// LS Electric XG5000 project: NewPLC
// PLC LSPLC
// module base 0 slot 0: 입력 모듈:XGI-D21A (DC 24V 입력, 8점 (전류소스/싱크입력))
// module base 0 slot 1: 입력 모듈:XGI-D22A/B (DC 24V 입력, 16점 (전류소스 싱크공용/ 전류소스 입력))
// module base 0 slot 2: 입력 모듈:XGI-D24A/B (DC 24V 입력, 32점 (전류소스 싱크공용/ 전류소스 입력))
// module base 0 slot 3: 입력 모듈:XGI-D28A/B (DC 24V 입력, 64점 (전류소스 싱크공용/ 전류소스 입력))
// module base 0 slot 4: 입력 모듈:XGI-A12A (AC 110V 입력, 16점)
// module base 0 slot 5: 입력 모듈:XGI-A21A/C (AC 220V 입력, 8점(8점/COM) / 8점(1점/COM))
// module base 0 slot 6: 입력 모듈:XGI-D21D (진단기능 내장형 DC24V 입력, 8점)
// module base 0 slot 7: 입출력 모듈:XGH-DT4A (DC 24V 입력, 트랜지스터 출력 32점 )
// module base 0 slot 8: 전용 모듈:XGI-LBDA (AC 110V 램프 단선검출 입력, 6점)
// module base 0 slot 9: 전용 모듈:XGI-LBDB (AC/DC 10V 램프 단선검출 입력, 6점)
// module base 0 slot 10: FDEnet:XGL-EDMT (전용 Ethernet 통신 모듈, 전기 Master)
// module base 0 slot 11: FDEnet:XGL-EDMF (전용 Ethernet 통신 모듈, 광 Master)
// module base 1 slot 0: 출력 모듈:XGQ-RY1A (릴레이 출력, 8점 (2A용, 단독 COM.))
// module base 1 slot 1: 출력 모듈:XGQ-RY2A/B (릴레이 출력, 16점 (2A용, Varistor 없음/Varistor 부착))
// module base 1 slot 2: 출력 모듈:XGQ-TR1C (트랜지스터 출력, 8점 (2A용, 싱크출력))
// module base 1 slot 3: 출력 모듈:XGQ-TR2A/B (트랜지스터 출력, 16점 (0.5A용, 싱크출력/소스출력))
// module base 1 slot 4: 출력 모듈:XGQ-TR4A/B (트랜지스터 출력, 32점 (0.1A용, 싱크출력/소스출력))
// module base 1 slot 5: 출력 모듈:XGQ-TR8A/B (트랜지스터 출력, 64점 (0.1A용, 싱크출력/소스출력))
// module base 1 slot 6: 출력 모듈:XGQ-SS2A (트라이액 출력, 16점 (1A용))
// module base 1 slot 7: 출력 모듈:XGQ-RY1D (진단기능 내장형 Relay 출력, 8점)
// module base 1 slot 8: 고속카운터 모듈:XGF-HO2A (고속카운터 펄스(OC) 입력형, 2채널)
// module base 1 slot 9: 고속카운터 모듈:XGF-HD2A (고속카운터 펄스(LD) 입력형, 2채널)
// module base 1 slot 10: 고속카운터 모듈:XGF-HO8A (고속카운터 펄스(OC) 입력형, 8채널)
// module base 1 slot 11: Dnet:XGL-DMEA/B (Dnet 통신 모듈, DeviceNet Master)
// module base 2 slot 0: 아날로그입력 모듈:XGF-AV8A (A/D 전압 입력형 8채널)
// module base 2 slot 1: 아날로그입력 모듈:XGF-AC8A (A/D 전류 입력형 8채널)
// module base 2 slot 2: 아날로그입력 모듈:XGF-AD4S (A/D 절연형 4채널)
// module base 2 slot 3: 아날로그입력 모듈:XGF-AD8A (A/D 전압/전류 입력형 8채널)
// module base 2 slot 4: 아날로그입력 모듈:XGF-AD16A (A/D 전압/전류 입력형 16채널)
// module base 2 slot 5: 아날로그입력 모듈:XGF-AC4H (HART 인터페이스 아날로그 전류입력, 4채널)
// module base 2 slot 6: 아날로그입력 모듈:XGF-AW4S (A/D 절연형 4채널(2선 입력형))
// module base 2 slot 7: 모션제어 모듈:XGF-M16M (모션 전용네트 (M-II)형, 16축)
// module base 2 slot 8: 모션제어 모듈:XGF-M32E (네트워크 표준형, 32축)
// module base 2 slot 9: 데이터로그 모듈:XGF-DL16A (데이터 로그 모듈)
// module base 2 slot 10: SOE모듈:XGF-SOEA (이벤트 기록 모듈)
// module base 2 slot 11: Rnet:XGL-RMEA/B (Rnet 통신 모듈, Rnet Master)
// module base 3 slot 0: 아날로그출력 모듈:XGF-DV4A (D/A 전압 출력형 4채널)
// module base 3 slot 1: 아날로그출력 모듈:XGF-DV8A (D/A 전압 출력형 8채널)
// module base 3 slot 2: 아날로그출력 모듈:XGF-DC4A (D/A 전류 출력형 4채널)
// module base 3 slot 3: 아날로그출력 모듈:XGF-DC8A (D/A 전류 출력형 8채널)
// module base 3 slot 4: 아날로그출력 모듈:XGF-DV4S (D/A 절연형 4채널(전압형))
// module base 3 slot 5: 아날로그출력 모듈:XGF-DC4S (D/A 절연형 4채널(전류형))
// module base 3 slot 6: 아날로그출력 모듈:XGF-DC4H (HART 인터페이스 아날로그 전류출력, 4채널)
// module base 3 slot 7: 아날로그출력 모듈:XGF-DA4S (D/A 절연형, 4채널)
// module base 3 slot 8: 온도입력 모듈:XGF-RD4A (온도 입력형 4채널)
// module base 3 slot 9: 온도입력 모듈:XGF-RD4S (온도 입력형 4채널(절연형))
// module base 3 slot 10: 온도입력 모듈:XGF-TC4S (온도 입력형 (절연형 4채널))
// module base 3 slot 11: 온도입력 모듈:XGF-RD8A (측온저항체 센서 입력형 8채널)

PROGRAM NewProgram (task: 스캔 프로그램)

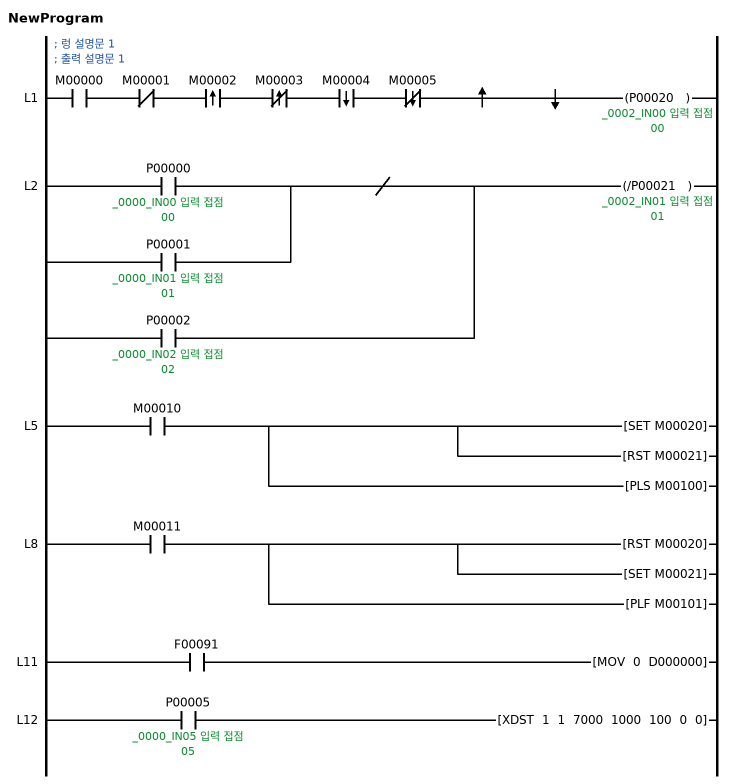
// 렁 설명문 1
; L1
LOAD      M00000
AND NOT   M00001
ANDP      M00002
ANDP NOT  M00003
ANDN      M00004
ANDN NOT  M00005
R_EDGE
F_EDGE
OUT       P00020	// _0002_IN00 입력 접점 00
// output comment: 출력 설명문 1
; L2
LOAD      P00000	// _0000_IN00 입력 접점 00
OR        P00001	// _0000_IN01 입력 접점 01
NOT
OR        P00002	// _0000_IN02 입력 접점 02
OUT NOT   P00021	// _0002_IN01 입력 접점 01
; L5
LOAD      M00010
SET       M00020
RST       M00021
OUTP      M00100
; L8
LOAD      M00011
RST       M00020
SET       M00021
OUTN      M00101
; L11
LOAD      F00091
MOV       0 D000000
; L12
LOAD      P00005	// _0000_IN05 입력 접점 05
XDST      1 1 7000 1000 100 0 0